FUNCTION_BLOCK FB_Buffer5 IMPLEMENTS ITF_Buffer5
VAR_INPUT
END_VAR
VAR_OUTPUT
END_VAR
VAR
END_VAR

{warning 'Add method implementation '}
METHOD Aborted : BOOL
END_METHOD

{warning 'Add method implementation '}
METHOD Aborting : BOOL
END_METHOD

{warning 'Add method implementation '}
METHOD Clearing : BOOL
END_METHOD

{warning 'Add method implementation '}
METHOD Execute : BOOL
END_METHOD

{warning 'Add method implementation '}
METHOD Held : BOOL
END_METHOD

{warning 'Add method implementation '}
METHOD Holding : BOOL
END_METHOD

{warning 'Add method implementation '}
METHOD Idle : BOOL
END_METHOD

{warning 'Add method implementation '}
METHOD Resetting : BOOL
END_METHOD

{warning 'Add method implementation '}
METHOD Starting : BOOL
END_METHOD

{warning 'Add method implementation '}
METHOD Stopped : BOOL
END_METHOD

{warning 'Add method implementation '}
METHOD Stopping : BOOL
END_METHOD

{warning 'Add method implementation '}
METHOD Suspended : BOOL
END_METHOD

{warning 'Add method implementation '}
METHOD Suspending : BOOL
END_METHOD

{warning 'Add method implementation '}
METHOD Unholding : BOOL
END_METHOD

{warning 'Add method implementation '}
METHOD Unsuspending : BOOL
END_METHOD

END_FUNCTION_BLOCK

(* stored: Version 1.1.0.1
   POU FB_Buffer5: Id {68b6c181-fb5e-4633-8340-2c972290f158}, SpecialFunc None
   Folder Methods: Id {ea3de5bf-78cc-4aaa-881d-872d01108b36}
   Method Aborted: Id {4d723c13-ef33-489d-93b0-ee0e47df53d1}
   Method Aborting: Id {e8243e2d-b98e-462f-aec6-a3e35b85de58}
   Method Clearing: Id {1ef713ba-ba14-4090-8697-df3273aa5286}
   Method Execute: Id {346565ed-a89d-4b29-b237-7f14c37fc0a3}
   Method Held: Id {1f68f14d-6aee-4cdb-b61c-3b93dbeddc9f}
   Method Holding: Id {2c6c7c69-5562-4745-8d05-7105f4ac9efc}
   Method Idle: Id {650c2b5e-fb8b-4b04-9c91-e984657e03bd}
   Method Resetting: Id {ef435268-8b2c-4149-8b13-5d991fe4e438}
   Method Starting: Id {fbdede14-24a4-48c5-a131-2bb90d797689}
   Method Stopped: Id {8c889838-6f6a-44b6-9deb-a2ed4be845af}
   Method Stopping: Id {22d11821-06b2-4886-8caf-a91b61c2870a}
   Method Suspended: Id {e6c5041e-6231-4110-9645-fbfc5a2a1797}
   Method Suspending: Id {f73956be-9c97-46b3-bd77-349510f69156}
   Method Unholding: Id {bd214273-4c3d-409e-bf69-3c9f96aacd9c}
   Method Unsuspending: Id {7d53bfdb-4229-44c8-8310-c79d7bc0b108} *)
